Fanuc KAREL source: kb00119.KL

-- PROVISIONAL review KL for V770-1; original PC SHA256 dbf07798081446707c5575ca28bd6f49ec1a97ceda8db5dd1be887101868e4c3
-- Incomplete behavior may be omitted. Consult companion uncertainty JSON. Do not deploy.
PROGRAM KB00119
%NOLOCKGROUP
BEGIN
  -- UNRESOLVED_PC offsets 5-12; opcodes 9D,23
  -- UNRESOLVED_PC offsets 17-24; opcodes 9D,23
  -- UNRESOLVED_PC offsets 29-45; opcodes 27,22,22,31
  -- UNRESOLVED_PC offsets 50-54; opcodes 7F
END KB00119
